(* Status of Stober PS6A34 *)

TYPE ST_STOEBER_PS6A34Status_1 :
STRUCT
	bReady				:BOOL;			(* Stoeber PS6A34 ready / StoeberPS6A34 i.O. *)
	bNoOverload			:BOOL;			(* StoeberPS6A34 no overload  / StoeberPS6A34 nicht überlastet *)
	bGridPhaseOk		:BOOL;			(* StoeberPS6A34 no grid phase failure  / StoeberPS6A34 nicht Netzphasenausfall *)
END_STRUCT
END_TYPE

(* stored: Version 1.1.0.1, ProductVersion 3.1.4024.15
   DUT ST_STOEBER_PS6A34Status_1: Id {087dd5c2-7fef-4d07-9bbc-17556b89dcc9} *)
